Fanuc KAREL source: KX00002.KL

PROGRAM KX00002
%NOLOCKGROUP
VAR
  I: INTEGER
  J: INTEGER
  B: BOOLEAN
  F: FILE
  S: STRING[80]
  P: XYZWPR
BEGIN
  OPEN FILE F ('RW', 'MD:KFSAMPLE.DT')
  CLOSE FILE F
END KX00002
